// TIA Portal V20 export
ORGANIZATION_BLOCK "OB1"   // OB1, STL, ProgramCycle
TITLE = "Main Program Sweep (Cycle)"
{ S7_Optimized_Access := 'FALSE' }
// stored: AutoNumber false
   VAR_TEMP
      OB1_EV_CLASS : Byte;   // Bits 0-3 = 1 (Coming event), Bits 4-7 = 1 (Event class 1)
      OB1_SCAN_1 : Byte;   // 1 (Cold restart scan 1 of OB 1), 3 (Scan 2-n of OB 1)
      OB1_PRIORITY : Byte;   // Priority of OB Execution
      OB1_OB_NUMBR : Byte;   // 1 (Organization block 1, OB1)
      OB1_RESERVED_1 : Byte;   // Reserved for system
      OB1_RESERVED_2 : Byte;   // Reserved for system
      OB1_PREV_CYCLE : Int;   // Cycle time of previous OB1 scan (milliseconds)
      OB1_MIN_CYCLE : Int;   // Minimum cycle time of OB1 (milliseconds)
      OB1_MAX_CYCLE : Int;   // Maximum cycle time of OB1 (milliseconds)
      OB1_DATE_TIME : Date_And_Time;   // Date and time OB1 started
   END_VAR
BEGIN

NETWORK
TITLE = IBS1 und IBS0 für Inbetriebnahmezwecke
      SET;
      =     "IBS1";

      CLR;
      =     "IBS0";


NETWORK
TITLE = Sicherheitstechnik
//  CALL  "01_FB_ Simulation", "01_FB_ Simulation_DB"// Simulation muss vor und nach der Sicherheitstechnik aufgerufen werden

      CALL  "DataFromSafey", "DataFromSafey_DB";
      CALL  "DataToSafety", "DataToSafety_DB";






NETWORK
TITLE = Allgemein



      CALL  "02_Wartungsfreigaben", "02_Wartungsfreigaben_DB";
      CALL  "03_Betriebsart", "03_Betriebsart_DB";


      CALL  "05_Not-Aus", "05_Not-Aus_DB";
      CALL  "06_Grundstellungen", "06_Grundstellungen_DB";




//     CALL  "01_FB_ Simulation", "01_FB_ Simulation_DB"// Simulation muss vor und nach der Sicherheitstechnik aufgerufen werden



NETWORK
TITLE = Zyklisch wechselnder Merker
      A     "Zyklisch wechselnder Merker";
      JC    M015;
      AN    "Zyklisch wechselnder Merker";
      S     "Zyklisch wechselnder Merker";
      JU    M016;
M015: NOP   0;
      R     "Zyklisch wechselnder Merker";
M016: NOP   0;


NETWORK
TITLE = 
      CALL  "Melden_VisuAllgemein", "Melden_VisuAllgemein_DB";
      CALL  "Schnittstelle SPS/HMI";
      CALL  "Störmeldungen";
      CALL  "Leuchtmelder Ampel", "Leuchtmelder Ampel_DB";


      CALL  "FB002_LabView", "DB002_LabView_DB";



      CALL  "Verwaltung_Teiledaten_FB", "Verwaltung_Teiledaten_FB_DB";

      CALL  "01_Alle_Zaehler", "01_Alle_Zaehler_DB";

      CALL  "02_Wartungszaehler", "02_Wartungszaehler_DB";


      CALL  "POS3_0_Bausteinaufrufe";


      CALL  "Zaehler_Sicherheit", "Zaehler_Sicherheit_DB";



NETWORK
TITLE = Simulation Eingänge in Zwischenspeicher sichern --> Muss im letzten Netzwerks stehen
//    CALL  MOVE
//         value_type:=Variant
//         IN  :="Simulation_DE200_bis_DE2199"
//         OUT :="01_FB_ Simulation_DB".DE200_bis_DE2199



END_ORGANIZATION_BLOCK
